INTERFACE ITcoRtc

PROPERTY IsSynchronized : BOOL
GET
END_GET
END_PROPERTY

PROPERTY IsValid : BOOL
GET
END_GET
END_PROPERTY

METHOD NowLocal : DATE_AND_TIME
END_METHOD

METHOD NowLocalAsTIMESTRUCT : Tc2_EtherCAT.Tc2_Utilities.TIMESTRUCT
END_METHOD

METHOD NowUTC : DATE_AND_TIME
END_METHOD

METHOD NowUTCAsTIMESTRUCT : Tc2_EtherCAT.Tc2_Utilities.TIMESTRUCT
END_METHOD

METHOD TickClock : ULINT
END_METHOD

END_INTERFACE

(* stored: Version 1.1.0.1
   Itf ITcoRtc: Id {f54bc528-8fdb-0177-2acd-c304b580985d}
   Property IsSynchronized: Id {e989db84-ead8-0485-3fa1-0445b66f52e3}
   Get Get: Id {3e920a2d-2ced-0e9d-3fe9-fcd40847fa88}
   Property IsValid: Id {66f4316f-7d87-0f76-192c-84fa99c1199a}
   Get Get: Id {e955570d-c675-0800-0743-44e0674472d7}
   Method NowLocal: Id {cb5c3e1b-5c35-049f-321a-41c43ce7891d}
   Method NowLocalAsTIMESTRUCT: Id {faf62912-5ac6-0765-13dd-eae44285ed7f}
   Method NowUTC: Id {66b88e73-4408-05c1-18eb-a65390fa484d}
   Method NowUTCAsTIMESTRUCT: Id {f75b99b9-fb58-07f6-0e63-76fe2d08bada}
   Method TickClock: Id {317ccaa2-fed5-0818-37bf-03f24bf02b0d} *)
